Fanuc KAREL source: KC00017.KL

PROGRAM KC00017
%NOLOCKGROUP
%ENVIRONMENT PBCORE
VAR
  I: INTEGER
  J: INTEGER
  K: INTEGER
  R: REAL
  B: BOOLEAN
  S: STRING[80]
  T: STRING[80]
  P: PATH
  Q: PATH
  AI: ARRAY[8] OF INTEGER
  AB: ARRAY[244] OF BYTE
  F: FILE
BEGIN
  READ_KB(F,S,I,J,K,I,T,I,J,K)
END KC00017
